(* PLC project PR_UnloadingSeq_Soft2.0_workflow_f29f28_PLC, SiemensToBackhoff Siemens TIA Portal → Beckhoff TwinCAT PLCopen Converter 2.2 *)
(* stored: creationDateTime 2026-10-12T09:25:58.949097, modificationDateTime 2026-10-12T09:25:58.949097 *)

FUNCTION_BLOCK PR_UnloadingSeq_Soft2.0_workflow_f29f28
VAR_INPUT
	iAbort : BOOL;
	iAutoRunning : BOOL;
	iFaultReset : BOOL;
	iGantryAtPick : BOOL;
	iManualEntryConfirm : BOOL;
	iPartPickOver : BOOL;
	iPartPresent : BOOL;
	iPickConfirmed : BOOL;
	iRFIDReadError : BOOL;
	iRFIDReadOver : BOOL;
	iRFWriteDone : BOOL;
	iRFWriteError : BOOL;
	iRTR_Frm_Gantry : BOOL;
	iReject : BOOL;
	iReset_fault : BOOL;
	iRetry : BOOL;
	iRetryCount : INT;
	iSstMode : BOOL;
	iSstPB : BOOL;
	iStartFrmFibroSeq : BOOL;
	iSystemAtHome : BOOL;
	iUnloadGantryAtSafe : BOOL;
END_VAR
VAR_OUTPUT
	qError : ARRAY[0..2] OF BOOL;
	qMessage : ARRAY[0..0] OF BOOL;
	qUnloadOver : BOOL;
END_VAR
VAR
	c120_ChkPartAbsent_T1 : BOOL;
	c120_ChkPartAbsent_T2 : BOOL;
	c130_WtOpDecisionPick_T1 : BOOL;
	c130_WtOpDecisionPick_T2 : BOOL;
	c140_WtRFIDWriteOver_T1 : BOOL;
	c140_WtRFIDWriteOver_T2 : BOOL;
	c150_ChkRFWriteRetryCount_T1 : BOOL;
	c150_ChkRFWriteRetryCount_T2 : BOOL;
	c160_WtOpDecisionWrite_T1 : BOOL;
	c160_WtOpDecisionWrite_T2 : BOOL;
	c20_ChkRecoveryStatus_T1 : BOOL;
	c20_ChkRecoveryStatus_T2 : BOOL;
	c20_ChkRecoveryStatus_T3 : BOOL;
	c50_WtRFIDReadOver_T1 : BOOL;
	c50_WtRFIDReadOver_T2 : BOOL;
	c60_ChkRetryCountOver_T1 : BOOL;
	c60_ChkRetryCountOver_T2 : BOOL;
	c70_WtOpDecisionRead_T1 : BOOL;
	c70_WtOpDecisionRead_T2 : BOOL;
	c80_ChkPartWorkable_T1 : BOOL;
	c80_ChkPartWorkable_T2 : BOOL;
	StateNo : INT;
	s100_WtGantryAtPick : BOOL;
	s100_WtGantryAtPick_T1 : BOOL;
	s10_WtStartFrmMain : BOOL;
	s10_WtStartFrmMain_T1 : BOOL;
	s110_WtPartPick : BOOL;
	s110_WtPartPick_T1 : BOOL;
	s120_ChkPartAbsent : BOOL;
	s120_ChkPartAbsent_T1 : BOOL;
	s120_ChkPartAbsent_T2 : BOOL;
	s130_WtOpDecisionPick : BOOL;
	s130_WtOpDecisionPick_T1 : BOOL;
	s130_WtOpDecisionPick_T2 : BOOL;
	s140_WtRFIDWriteOver : BOOL;
	s140_WtRFIDWriteOver_T1 : BOOL;
	s140_WtRFIDWriteOver_T2 : BOOL;
	s150_ChkRFWriteRetryCount : BOOL;
	s150_ChkRFWriteRetryCount_T1 : BOOL;
	s150_ChkRFWriteRetryCount_T2 : BOOL;
	s160_WtOpDecisionWrite : BOOL;
	s160_WtOpDecisionWrite_T1 : BOOL;
	s160_WtOpDecisionWrite_T2 : BOOL;
	s170_ChkSystemAtHome : BOOL;
	s170_ChkSystemAtHome_T1 : BOOL;
	s180_WtStartLow : BOOL;
	s180_WtStartLow_T1 : BOOL;
	s1_WtResetReleased : BOOL;
	s1_WtResetReleased_T1 : BOOL;
	s20_ChkRecoveryStatus : BOOL;
	s20_ChkRecoveryStatus_T1 : BOOL;
	s20_ChkRecoveryStatus_T2 : BOOL;
	s20_ChkRecoveryStatus_T3 : BOOL;
	s30_WtOperatorAck : BOOL;
	s30_WtOperatorAck_T1 : BOOL;
	s40_WtAllAxesSafe : BOOL;
	s40_WtAllAxesSafe_T1 : BOOL;
	s50_WtRFIDReadOver : BOOL;
	s50_WtRFIDReadOver_T1 : BOOL;
	s50_WtRFIDReadOver_T2 : BOOL;
	s60_ChkRetryCountOver : BOOL;
	s60_ChkRetryCountOver_T1 : BOOL;
	s60_ChkRetryCountOver_T2 : BOOL;
	s70_WtOpDecisionRead : BOOL;
	s70_WtOpDecisionRead_T1 : BOOL;
	s70_WtOpDecisionRead_T2 : BOOL;
	s80_ChkPartWorkable : BOOL;
	s80_ChkPartWorkable_T1 : BOOL;
	s80_ChkPartWorkable_T2 : BOOL;
	s90_WtRTRFrmGantry : BOOL;
	s90_WtRTRFrmGantry_T1 : BOOL;
	sAbnormalStatus : BOOL;
	sPartWorkable : BOOL;
	sRFReadRetryCount : INT;
	sRFWriteRetryCount : INT;
	sSst : BOOL;
	sSstPulse : BOOL;
	sSstRise : R_TRIG;
	sStWtResetRel : BOOL;
	sStWtResetRel_T1 : BOOL;
	sUnloadingActive : BOOL;
END_VAR
VAR_TEMP
	tOne : BOOL;
END_VAR
  VAR  (* added by the conversion: wires and edge detectors of the diagram *)
    _w24 : BOOL;
    _w26 : BOOL;
    _w39 : BOOL;
    _w41 : BOOL;
    _w42 : BOOL;
    _w59 : BOOL;
    _w61 : BOOL;
    _w62 : BOOL;
    _w95 : BOOL;
    _w99 : BOOL;
    _w100 : BOOL;
    _w101 : BOOL;
    _w102 : BOOL;
    _w115 : BOOL;
    _w117 : BOOL;
    _w118 : BOOL;
    _w135 : BOOL;
    _w137 : BOOL;
    _w138 : BOOL;
    _w162 : BOOL;
    _w166 : BOOL;
    _w167 : BOOL;
    _w168 : BOOL;
    _w202 : BOOL;
    _w204 : BOOL;
    _w205 : BOOL;
    _w206 : BOOL;
    _w230 : BOOL;
    _w232 : BOOL;
    _w233 : BOOL;
    _w234 : BOOL;
    _w262 : BOOL;
    _w265 : BOOL;
    _w266 : BOOL;
    _w267 : BOOL;
    _w280 : BOOL;
    _w283 : BOOL;
    _w284 : BOOL;
    _w297 : BOOL;
    _w300 : BOOL;
    _w301 : BOOL;
    _w314 : BOOL;
    _w317 : BOOL;
    _w318 : BOOL;
    _w343 : BOOL;
    _w345 : BOOL;
    _w346 : BOOL;
    _w347 : BOOL;
    _w371 : BOOL;
    _w373 : BOOL;
    _w374 : BOOL;
    _w375 : BOOL;
    _w399 : BOOL;
    _w404 : BOOL;
    _w405 : BOOL;
    _w406 : BOOL;
    _w440 : BOOL;
    _w442 : BOOL;
    _w443 : BOOL;
    _w444 : BOOL;
    _w469 : BOOL;
    _w471 : BOOL;
    _w472 : BOOL;
    _w473 : BOOL;
    _w495 : BOOL;
    _w498 : BOOL;
    _w499 : BOOL;
    _w517 : BOOL;
    _w519 : BOOL;
    _w520 : BOOL;
  END_VAR

(* LD diagram, written out as Structured Text *)
(* Network 1 *)
(* Create Single Step Pulse bit *)
(* Create Single Step bit *)
(* Transition for STATE Num:0 Reset Released *)
(* STATE Num:0 Reset Released *)
(* Transition for STATE Num:1 Wait For Reset Released *)
(* STATE Num:1 Wait For Reset Released *)
(* Transition for STATE Num:10 Wait for Start from Main Sequence *)
(* STATE Num:10 Wait for Start from Main Sequence *)
(* Condition1 for STATE Num:20 Chek Recovery Status *)
(* Condition2 for STATE Num:20 Chek Recovery Status *)
(* Condition3 for STATE Num:20 Chek Recovery Status *)
(* Transition for STATE Num:20 Chek Recovery Status *)
(* STATE Num:20 Chek Recovery Status *)
(* Transition for STATE Num:30 Wait for Operator Ack *)
(* STATE Num:30 Wait for Operator Ack *)
(* Actions for STATE Num:30 Wait for Operator Ack *)
(* Transition for STATE Num:40 Wait For All Axes are Safe *)
(* STATE Num:40 Wait For All Axes are Safe *)
(* Condition1 for STATE Num:50 Wait For RFID Read Over *)
(* Condition2 for STATE Num:50 Wait For RFID Read Over *)
(* Transition for STATE Num:50 Wait For RFID Read Over *)
(* STATE Num:50 Wait For RFID Read Over *)
(* Transition Action for STATE Num:50 Condition1 increment sRFReadRetryCount *)
(* Condition1 for STATE Num:60 Check Retry Count Over *)
(* Condition2 for STATE Num:60 Check Retry Count Over *)
(* Transition for STATE Num:60 Check Retry Count Over *)
(* STATE Num:60 Check Retry Count Over *)
(* Condition1 for STATE Num:70 Wait For Operator Decision_Read *)
(* Condition2 for STATE Num:70 Wait For Operator Decision_Read *)
(* Transition for STATE Num:70 Wait For Operator Decision_Read *)
(* STATE Num:70 Wait For Operator Decision_Read *)
(* Actions for STATE Num:70 Wait For Operator Decision_Read *)
(* Condition1 for STATE Num:80 Check Part is Workable *)
(* Condition2 for STATE Num:80 Check Part is Workable *)
(* Transition for STATE Num:80 Check Part is Workable *)
(* STATE Num:80 Check Part is Workable *)
(* Transition for STATE Num:90 Wait For RTR From Unload gantry *)
(* STATE Num:90 Wait For RTR From Unload gantry *)
(* Transition for STATE Num:100 Wait Gantry at Pick Position *)
(* STATE Num:100 Wait Gantry at Pick Position *)
(* Transition for STATE Num:110 Wait For Part Pick *)
(* STATE Num:110 Wait For Part Pick *)
(* Condition1 for STATE Num:120 Check Part Absent *)
(* Condition2 for STATE Num:120 Check Part Absent *)
(* Transition for STATE Num:120 Check Part Absent *)
(* STATE Num:120 Check Part Absent *)
(* Condition1 for STATE Num:130 Wait For Operator Decision_Pick *)
(* Condition2 for STATE Num:130 Wait For Operator Decision_Pick *)
(* Transition for STATE Num:130 Wait For Operator Decision_Pick *)
(* STATE Num:130 Wait For Operator Decision_Pick *)
(* Condition1 for STATE Num:140 Wait for RFID Write Over *)
(* Condition2 for STATE Num:140 Wait for RFID Write Over *)
(* Transition for STATE Num:140 Wait for RFID Write Over *)
(* STATE Num:140 Wait for RFID Write Over *)
(* Transition Action for STATE Num:140 Condition1 increment sRFWriteRetryCount *)
(* Condition1 for STATE Num:150 Check RFID Write Retry Count Over *)
(* Condition2 for STATE Num:150 Check RFID Write Retry Count Over *)
(* Transition for STATE Num:150 Check RFID Write Retry Count Over *)
(* STATE Num:150 Check RFID Write Retry Count Over *)
(* Condition1 for STATE Num:160 Wait For Operator Decision_Write *)
(* Condition2 for STATE Num:160 Wait For Operator Decision_Write *)
(* Transition for STATE Num:160 Wait For Operator Decision_Write *)
(* STATE Num:160 Wait For Operator Decision_Write *)
(* Transition Action for STATE Num:160 Condition1 set qError2 and qMessage0 *)
(* Transition Action for STATE Num:160 Condition2 set qError2 *)
(* Transition for STATE Num:170 Check System at Home_Safe for Index *)
(* STATE Num:170 Check System at Home_Safe for Index *)
(* Transition for STATE Num:180 Wait for Start Low *)
(* STATE Num:180 Wait for Start Low *)
tOne := tOne OR NOT tOne;
sSstRise(CLK := iSstPB);
sSstPulse := sSstRise.Q;
sSst := iSstMode AND sSstPulse OR NOT iSstMode;
sStWtResetRel_T1 := sStWtResetRel AND iAutoRunning;
_w24 := sStWtResetRel;
_w26 := (_w24 OR NOT iAutoRunning) AND NOT sStWtResetRel_T1;
sStWtResetRel := _w26;
IF _w26 THEN StateNo := 0; END_IF;
s1_WtResetReleased_T1 := s1_WtResetReleased AND NOT sStWtResetRel AND sSst AND iAutoRunning;
_w39 := s1_WtResetReleased;
_w41 := (_w39 OR sStWtResetRel_T1) AND NOT sStWtResetRel;
_w42 := _w41 AND NOT s1_WtResetReleased_T1;
s1_WtResetReleased := _w42;
IF _w42 THEN StateNo := 1; END_IF;
s10_WtStartFrmMain_T1 := s10_WtStartFrmMain AND NOT sStWtResetRel AND sSst AND iStartFrmFibroSeq;
IF s10_WtStartFrmMain AND NOT sStWtResetRel AND sSst AND iStartFrmFibroSeq THEN sRFReadRetryCount := 0; END_IF;
IF s10_WtStartFrmMain AND NOT sStWtResetRel AND sSst AND iStartFrmFibroSeq THEN sRFWriteRetryCount := 0; END_IF;
_w59 := s10_WtStartFrmMain;
_w61 := (_w59 OR s1_WtResetReleased_T1) AND NOT sStWtResetRel;
_w62 := _w61 AND NOT s10_WtStartFrmMain_T1;
s10_WtStartFrmMain := _w62;
IF _w62 THEN StateNo := 10; END_IF;
c20_ChkRecoveryStatus_T1 := sAbnormalStatus;
c20_ChkRecoveryStatus_T2 := sUnloadingActive;
c20_ChkRecoveryStatus_T3 := NOT sAbnormalStatus AND NOT sUnloadingActive;
s20_ChkRecoveryStatus_T1 := s20_ChkRecoveryStatus AND NOT sStWtResetRel AND sSst AND c20_ChkRecoveryStatus_T1;
s20_ChkRecoveryStatus_T2 := s20_ChkRecoveryStatus AND NOT sStWtResetRel AND sSst AND NOT s20_ChkRecoveryStatus_T1 AND c20_ChkRecoveryStatus_T2;
s20_ChkRecoveryStatus_T3 := s20_ChkRecoveryStatus AND NOT sStWtResetRel AND sSst AND NOT s20_ChkRecoveryStatus_T1 AND NOT s20_ChkRecoveryStatus_T1 AND NOT s20_ChkRecoveryStatus_T2 AND c20_ChkRecoveryStatus_T3;
_w95 := s20_ChkRecoveryStatus;
_w99 := (_w95 OR s10_WtStartFrmMain_T1 OR s30_WtOperatorAck_T1 OR s180_WtStartLow_T1) AND NOT sStWtResetRel;
_w100 := _w99 AND NOT s20_ChkRecoveryStatus_T1;
_w101 := _w100 AND NOT s20_ChkRecoveryStatus_T2;
_w102 := _w101 AND NOT s20_ChkRecoveryStatus_T3;
s20_ChkRecoveryStatus := _w102;
IF _w102 THEN StateNo := 20; END_IF;
s30_WtOperatorAck_T1 := s30_WtOperatorAck AND NOT sStWtResetRel AND sSst AND iFaultReset;
_w115 := s30_WtOperatorAck;
_w117 := (_w115 OR s20_ChkRecoveryStatus_T1) AND NOT sStWtResetRel;
_w118 := _w117 AND NOT s30_WtOperatorAck_T1;
s30_WtOperatorAck := _w118;
IF _w118 THEN StateNo := 30; END_IF;
qError[0] := s30_WtOperatorAck;
s40_WtAllAxesSafe_T1 := s40_WtAllAxesSafe AND NOT sStWtResetRel AND sSst AND iUnloadGantryAtSafe;
_w135 := s40_WtAllAxesSafe;
_w137 := (_w135 OR s20_ChkRecoveryStatus_T3) AND NOT sStWtResetRel;
_w138 := _w137 AND NOT s40_WtAllAxesSafe_T1;
s40_WtAllAxesSafe := _w138;
IF _w138 THEN StateNo := 40; END_IF;
c50_WtRFIDReadOver_T1 := iRFIDReadError;
c50_WtRFIDReadOver_T2 := iRFIDReadOver;
s50_WtRFIDReadOver_T1 := s50_WtRFIDReadOver AND NOT sStWtResetRel AND sSst AND c50_WtRFIDReadOver_T1;
s50_WtRFIDReadOver_T2 := s50_WtRFIDReadOver AND NOT sStWtResetRel AND sSst AND NOT s50_WtRFIDReadOver_T1 AND c50_WtRFIDReadOver_T2;
_w162 := s50_WtRFIDReadOver;
_w166 := (_w162 OR s40_WtAllAxesSafe_T1 OR s60_ChkRetryCountOver_T2 OR s70_WtOpDecisionRead_T1) AND NOT sStWtResetRel;
_w167 := _w166 AND NOT s50_WtRFIDReadOver_T1;
_w168 := _w167 AND NOT s50_WtRFIDReadOver_T2;
s50_WtRFIDReadOver := _w168;
IF _w168 THEN StateNo := 50; END_IF;
IF s50_WtRFIDReadOver_T1 THEN sRFReadRetryCount := sRFReadRetryCount + 1; END_IF;
c60_ChkRetryCountOver_T1 := sRFReadRetryCount > iRetryCount;
c60_ChkRetryCountOver_T2 := sRFReadRetryCount <= iRetryCount;
s60_ChkRetryCountOver_T1 := s60_ChkRetryCountOver AND NOT sStWtResetRel AND sSst AND c60_ChkRetryCountOver_T1;
s60_ChkRetryCountOver_T2 := s60_ChkRetryCountOver AND NOT sStWtResetRel AND sSst AND NOT s60_ChkRetryCountOver_T1 AND c60_ChkRetryCountOver_T2;
_w202 := s60_ChkRetryCountOver;
_w204 := (_w202 OR s50_WtRFIDReadOver_T1) AND NOT sStWtResetRel;
_w205 := _w204 AND NOT s60_ChkRetryCountOver_T1;
_w206 := _w205 AND NOT s60_ChkRetryCountOver_T2;
s60_ChkRetryCountOver := _w206;
IF _w206 THEN StateNo := 60; END_IF;
c70_WtOpDecisionRead_T1 := iRetry;
c70_WtOpDecisionRead_T2 := iManualEntryConfirm;
s70_WtOpDecisionRead_T1 := s70_WtOpDecisionRead AND NOT sStWtResetRel AND sSst AND c70_WtOpDecisionRead_T1;
s70_WtOpDecisionRead_T2 := s70_WtOpDecisionRead AND NOT sStWtResetRel AND sSst AND NOT s70_WtOpDecisionRead_T1 AND c70_WtOpDecisionRead_T2;
_w230 := s70_WtOpDecisionRead;
_w232 := (_w230 OR s60_ChkRetryCountOver_T1) AND NOT sStWtResetRel;
_w233 := _w232 AND NOT s70_WtOpDecisionRead_T1;
_w234 := _w233 AND NOT s70_WtOpDecisionRead_T2;
s70_WtOpDecisionRead := _w234;
IF _w234 THEN StateNo := 70; END_IF;
qError[1] := s70_WtOpDecisionRead;
c80_ChkPartWorkable_T1 := NOT sPartWorkable;
c80_ChkPartWorkable_T2 := sPartWorkable;
s80_ChkPartWorkable_T1 := s80_ChkPartWorkable AND NOT sStWtResetRel AND sSst AND c80_ChkPartWorkable_T1;
s80_ChkPartWorkable_T2 := s80_ChkPartWorkable AND NOT sStWtResetRel AND sSst AND NOT s80_ChkPartWorkable_T1 AND c80_ChkPartWorkable_T2;
_w262 := s80_ChkPartWorkable;
_w265 := (_w262 OR s50_WtRFIDReadOver_T2 OR s70_WtOpDecisionRead_T2) AND NOT sStWtResetRel;
_w266 := _w265 AND NOT s80_ChkPartWorkable_T1;
_w267 := _w266 AND NOT s80_ChkPartWorkable_T2;
s80_ChkPartWorkable := _w267;
IF _w267 THEN StateNo := 80; END_IF;
s90_WtRTRFrmGantry_T1 := s90_WtRTRFrmGantry AND NOT sStWtResetRel AND sSst AND iRTR_Frm_Gantry;
_w280 := s90_WtRTRFrmGantry;
_w283 := (_w280 OR s80_ChkPartWorkable_T1 OR s80_ChkPartWorkable_T2) AND NOT sStWtResetRel;
_w284 := _w283 AND NOT s90_WtRTRFrmGantry_T1;
s90_WtRTRFrmGantry := _w284;
IF _w284 THEN StateNo := 90; END_IF;
s100_WtGantryAtPick_T1 := s100_WtGantryAtPick AND NOT sStWtResetRel AND sSst AND iGantryAtPick;
_w297 := s100_WtGantryAtPick;
_w300 := (_w297 OR s90_WtRTRFrmGantry_T1 OR s130_WtOpDecisionPick_T1) AND NOT sStWtResetRel;
_w301 := _w300 AND NOT s100_WtGantryAtPick_T1;
s100_WtGantryAtPick := _w301;
IF _w301 THEN StateNo := 100; END_IF;
s110_WtPartPick_T1 := s110_WtPartPick AND NOT sStWtResetRel AND sSst AND iPartPickOver;
_w314 := s110_WtPartPick;
_w317 := (_w314 OR s100_WtGantryAtPick_T1 OR s20_ChkRecoveryStatus_T2) AND NOT sStWtResetRel;
_w318 := _w317 AND NOT s110_WtPartPick_T1;
s110_WtPartPick := _w318;
sUnloadingActive := _w318;
IF _w318 THEN StateNo := 110; END_IF;
c120_ChkPartAbsent_T1 := iPartPresent;
c120_ChkPartAbsent_T2 := NOT iPartPresent;
s120_ChkPartAbsent_T1 := s120_ChkPartAbsent AND NOT sStWtResetRel AND sSst AND c120_ChkPartAbsent_T1;
s120_ChkPartAbsent_T2 := s120_ChkPartAbsent AND NOT sStWtResetRel AND sSst AND NOT s120_ChkPartAbsent_T1 AND c120_ChkPartAbsent_T2;
_w343 := s120_ChkPartAbsent;
_w345 := (_w343 OR s110_WtPartPick_T1) AND NOT sStWtResetRel;
_w346 := _w345 AND NOT s120_ChkPartAbsent_T1;
_w347 := _w346 AND NOT s120_ChkPartAbsent_T2;
s120_ChkPartAbsent := _w347;
IF _w347 THEN StateNo := 120; END_IF;
c130_WtOpDecisionPick_T1 := iRetry;
c130_WtOpDecisionPick_T2 := iPickConfirmed;
s130_WtOpDecisionPick_T1 := s130_WtOpDecisionPick AND NOT sStWtResetRel AND sSst AND c130_WtOpDecisionPick_T1;
s130_WtOpDecisionPick_T2 := s130_WtOpDecisionPick AND NOT sStWtResetRel AND sSst AND NOT s130_WtOpDecisionPick_T1 AND c130_WtOpDecisionPick_T2;
_w371 := s130_WtOpDecisionPick;
_w373 := (_w371 OR s120_ChkPartAbsent_T1) AND NOT sStWtResetRel;
_w374 := _w373 AND NOT s130_WtOpDecisionPick_T1;
_w375 := _w374 AND NOT s130_WtOpDecisionPick_T2;
s130_WtOpDecisionPick := _w375;
IF _w375 THEN StateNo := 130; END_IF;
c140_WtRFIDWriteOver_T1 := iRFWriteError;
c140_WtRFIDWriteOver_T2 := iRFWriteDone;
s140_WtRFIDWriteOver_T1 := s140_WtRFIDWriteOver AND NOT sStWtResetRel AND sSst AND c140_WtRFIDWriteOver_T1;
s140_WtRFIDWriteOver_T2 := s140_WtRFIDWriteOver AND NOT sStWtResetRel AND sSst AND NOT s140_WtRFIDWriteOver_T1 AND c140_WtRFIDWriteOver_T2;
_w399 := s140_WtRFIDWriteOver;
_w404 := (_w399 OR s120_ChkPartAbsent_T2 OR s130_WtOpDecisionPick_T2 OR s150_ChkRFWriteRetryCount_T2 OR s160_WtOpDecisionWrite_T2) AND NOT sStWtResetRel;
_w405 := _w404 AND NOT s140_WtRFIDWriteOver_T1;
_w406 := _w405 AND NOT s140_WtRFIDWriteOver_T2;
s140_WtRFIDWriteOver := _w406;
IF _w406 THEN StateNo := 140; END_IF;
IF s140_WtRFIDWriteOver_T1 THEN sRFWriteRetryCount := sRFWriteRetryCount + 1; END_IF;
c150_ChkRFWriteRetryCount_T1 := sRFWriteRetryCount > iRetryCount;
c150_ChkRFWriteRetryCount_T2 := sRFWriteRetryCount <= iRetryCount;
s150_ChkRFWriteRetryCount_T1 := s150_ChkRFWriteRetryCount AND NOT sStWtResetRel AND sSst AND c150_ChkRFWriteRetryCount_T1;
s150_ChkRFWriteRetryCount_T2 := s150_ChkRFWriteRetryCount AND NOT sStWtResetRel AND sSst AND NOT s150_ChkRFWriteRetryCount_T1 AND c150_ChkRFWriteRetryCount_T2;
_w440 := s150_ChkRFWriteRetryCount;
_w442 := (_w440 OR s140_WtRFIDWriteOver_T1) AND NOT sStWtResetRel;
_w443 := _w442 AND NOT s150_ChkRFWriteRetryCount_T1;
_w444 := _w443 AND NOT s150_ChkRFWriteRetryCount_T2;
s150_ChkRFWriteRetryCount := _w444;
IF _w444 THEN StateNo := 150; END_IF;
c160_WtOpDecisionWrite_T1 := iAbort OR iReject;
c160_WtOpDecisionWrite_T2 := iRetry;
s160_WtOpDecisionWrite_T1 := s160_WtOpDecisionWrite AND NOT sStWtResetRel AND sSst AND c160_WtOpDecisionWrite_T1;
s160_WtOpDecisionWrite_T2 := s160_WtOpDecisionWrite AND NOT sStWtResetRel AND sSst AND NOT s160_WtOpDecisionWrite_T1 AND c160_WtOpDecisionWrite_T2;
_w469 := s160_WtOpDecisionWrite;
_w471 := (_w469 OR s150_ChkRFWriteRetryCount_T1) AND NOT sStWtResetRel;
_w472 := _w471 AND NOT s160_WtOpDecisionWrite_T1;
_w473 := _w472 AND NOT s160_WtOpDecisionWrite_T2;
s160_WtOpDecisionWrite := _w473;
IF _w473 THEN StateNo := 160; END_IF;
qError[2] := s160_WtOpDecisionWrite_T1;
qMessage[0] := s160_WtOpDecisionWrite_T1;
qError[2] := s160_WtOpDecisionWrite_T2;
s170_ChkSystemAtHome_T1 := s170_ChkSystemAtHome AND NOT sStWtResetRel AND sSst AND iSystemAtHome;
_w495 := s170_ChkSystemAtHome;
_w498 := (_w495 OR s140_WtRFIDWriteOver_T2 OR s160_WtOpDecisionWrite_T1) AND NOT sStWtResetRel;
_w499 := _w498 AND NOT s170_ChkSystemAtHome_T1;
s170_ChkSystemAtHome := _w499;
IF _w499 THEN StateNo := 170; END_IF;
s180_WtStartLow_T1 := s180_WtStartLow AND NOT sStWtResetRel AND sSst AND NOT iStartFrmFibroSeq;
IF s180_WtStartLow AND NOT sStWtResetRel AND sSst AND NOT iStartFrmFibroSeq THEN sUnloadingActive := FALSE; END_IF;
IF s180_WtStartLow AND NOT sStWtResetRel AND sSst AND NOT iStartFrmFibroSeq THEN sRFReadRetryCount := 0; END_IF;
IF s180_WtStartLow AND NOT sStWtResetRel AND sSst AND NOT iStartFrmFibroSeq THEN sRFWriteRetryCount := 0; END_IF;
_w517 := s180_WtStartLow;
_w519 := (_w517 OR s170_ChkSystemAtHome_T1) AND NOT sStWtResetRel;
_w520 := _w519 AND NOT s180_WtStartLow_T1;
s180_WtStartLow := _w520;
IF _w520 THEN StateNo := 180; END_IF;
END_FUNCTION_BLOCK
